(* PLC project GeneratedProgram, SafePLC-Gen SafePLC-Gen Multimodal 1.0 *)
(* stored: creationDateTime 2026-04-25T12:02:49.071447Z *)

PROGRAM GeneratedProgram
  VAR
    FirstScan : BOOL;
    TI_2909_Scaled : REAL;
    TT_2909_Scaled : REAL;
    TT_2911_Scaled : REAL;
    TT_2917_Scaled : REAL;
    TI_2917_Scaled : REAL;
    XI_2901A_Scaled : REAL;
    XI_2901B_Scaled : REAL;
    TI_2909_HH_SP : REAL;
    TI_2909_H_SP : REAL;
    TI_2909_L_SP : REAL;
    TI_2909_LL_SP : REAL;
    TI_2909_Deadband : REAL;
    TI_2909_HH_Latch : BOOL;
    TI_2909_LL_Latch : BOOL;
    TI_2909_HH : BOOL;
    TI_2909_H : BOOL;
    TI_2909_L : BOOL;
    TI_2909_LL : BOOL;
    TI_2909_HH_Ack : BOOL;
    TI_2909_LL_Ack : BOOL;
    TT_2909_HH_SP : REAL;
    TT_2909_H_SP : REAL;
    TT_2909_L_SP : REAL;
    TT_2909_LL_SP : REAL;
    TT_2909_Deadband : REAL;
    TT_2909_HH_Latch : BOOL;
    TT_2909_LL_Latch : BOOL;
    TT_2909_HH : BOOL;
    TT_2909_H : BOOL;
    TT_2909_L : BOOL;
    TT_2909_LL : BOOL;
    TT_2909_HH_Ack : BOOL;
    TT_2909_LL_Ack : BOOL;
    TT_2911_HH_SP : REAL;
    TT_2911_H_SP : REAL;
    TT_2911_L_SP : REAL;
    TT_2911_LL_SP : REAL;
    TT_2911_Deadband : REAL;
    TT_2911_HH_Latch : BOOL;
    TT_2911_LL_Latch : BOOL;
    TT_2911_HH : BOOL;
    TT_2911_H : BOOL;
    TT_2911_L : BOOL;
    TT_2911_LL : BOOL;
    TT_2911_HH_Ack : BOOL;
    TT_2911_LL_Ack : BOOL;
    TT_2917_HH_SP : REAL;
    TT_2917_H_SP : REAL;
    TT_2917_L_SP : REAL;
    TT_2917_LL_SP : REAL;
    TT_2917_Deadband : REAL;
    TT_2917_HH_Latch : BOOL;
    TT_2917_LL_Latch : BOOL;
    TT_2917_HH : BOOL;
    TT_2917_H : BOOL;
    TT_2917_L : BOOL;
    TT_2917_LL : BOOL;
    TT_2917_HH_Ack : BOOL;
    TT_2917_LL_Ack : BOOL;
    TI_2917_HH_SP : REAL;
    TI_2917_H_SP : REAL;
    TI_2917_L_SP : REAL;
    TI_2917_LL_SP : REAL;
    TI_2917_Deadband : REAL;
    TI_2917_HH_Latch : BOOL;
    TI_2917_LL_Latch : BOOL;
    TI_2917_HH : BOOL;
    TI_2917_H : BOOL;
    TI_2917_L : BOOL;
    TI_2917_LL : BOOL;
    TI_2917_HH_Ack : BOOL;
    TI_2917_LL_Ack : BOOL;
    XI_2901A_HH_SP : REAL;
    XI_2901A_H_SP : REAL;
    XI_2901A_L_SP : REAL;
    XI_2901A_LL_SP : REAL;
    XI_2901A_Deadband : REAL;
    XI_2901A_HH_Latch : BOOL;
    XI_2901A_LL_Latch : BOOL;
    XI_2901A_HH : BOOL;
    XI_2901A_H : BOOL;
    XI_2901A_L : BOOL;
    XI_2901A_LL : BOOL;
    XI_2901A_HH_Ack : BOOL;
    XI_2901A_LL_Ack : BOOL;
    XI_2901B_HH_SP : REAL;
    XI_2901B_H_SP : REAL;
    XI_2901B_L_SP : REAL;
    XI_2901B_LL_SP : REAL;
    XI_2901B_Deadband : REAL;
    XI_2901B_HH_Latch : BOOL;
    XI_2901B_LL_Latch : BOOL;
    XI_2901B_HH : BOOL;
    XI_2901B_H : BOOL;
    XI_2901B_L : BOOL;
    XI_2901B_LL : BOOL;
    XI_2901B_HH_Ack : BOOL;
    XI_2901B_LL_Ack : BOOL;
    LOOP_2917_TRIP : BOOL;
    LOOP_2901A_TRIP : BOOL;
    LOOP_2901B_TRIP : BOOL;
    VSHH_2901A_HH : BOOL;
    VSHH_2901A_LL : BOOL;
    VSHH_2901B_HH : BOOL;
    VSHH_2901B_LL : BOOL;
    SAFE_STATE : BOOL;
    MCC_A_Run : BOOL;
    MCC_B_Run : BOOL;
    MCC_A_Out : BOOL;
    MCC_B_Out : BOOL;
    Drive_A_SP : REAL;
    Drive_B_SP : REAL;
    Drive_A_Kp : REAL;
    Drive_A_Ki : REAL;
    Drive_B_Kp : REAL;
    Drive_B_Ki : REAL;
    Drive_A_Error : REAL;
    Drive_B_Error : REAL;
    Drive_A_Integral : REAL;
    Drive_B_Integral : REAL;
    Drive_A_Output : REAL;
    Drive_B_Output : REAL;
    StartDelay_A : TON;
    StartDelay_B : TON;
    RS_2901_Inlet_A_Upper : BOOL;
    RS_2901_Inlet_A_Lower : BOOL;
    RS_2901_Outlet_B_Upper : BOOL;
    RS_2901_Outlet_B_Lower : BOOL;
    BV_Inlet_A_Upper_1 : BOOL;
    BV_Inlet_A_Upper_2 : BOOL;
    BV_Inlet_A_Lower_1 : BOOL;
    BV_Inlet_A_Lower_2 : BOOL;
    BV_Outlet_B_Upper_1 : BOOL;
    BV_Outlet_B_Upper_2 : BOOL;
    BV_Outlet_B_Lower_1 : BOOL;
    BV_Outlet_B_Lower_2 : BOOL;
    CV_HY_2903A_1 : BOOL;
    CV_HY_2903A_2 : BOOL;
    CV_HY_2903B_1 : BOOL;
    CV_HY_2903B_2 : BOOL;
    CSO_Inlet_1 : BOOL;
    CSO_Inlet_2 : BOOL;
    FLV_Inlet : BOOL;
    BV_1IN_Drain : BOOL;
    Breather_A_8IN : BOOL;
    Breather_B_8IN : BOOL;
    NC_Valve_Outlet : BOOL;
    System_Alarm : BOOL;
  END_VAR

            IF FirstScan THEN
    LOOP_2917_TRIP          := TRUE;
    LOOP_2901A_TRIP         := TRUE;
    LOOP_2901B_TRIP         := TRUE;
    SAFE_STATE              := TRUE;
    MCC_A_Out               := FALSE;
    MCC_B_Out               := FALSE;
    MCC_A_Run               := FALSE;
    MCC_B_Run               := FALSE;
    HY_2903A_Out            := 6554;
    HY_2903B_Out            := 6554;
    KV_2904                 := FALSE;
    XL_2901A                := FALSE;
    XL_2901B                := FALSE;
    XA_2901A                := FALSE;
    XA_2901B                := FALSE;
    TI_2909_HH_Latch        := FALSE;
    TI_2909_LL_Latch        := FALSE;
    TT_2909_HH_Latch        := FALSE;
    TT_2909_LL_Latch        := FALSE;
    TT_2911_HH_Latch        := FALSE;
    TT_2911_LL_Latch        := FALSE;
    TT_2917_HH_Latch        := FALSE;
    TT_2917_LL_Latch        := FALSE;
    TI_2917_HH_Latch        := FALSE;
    TI_2917_LL_Latch        := FALSE;
    XI_2901A_HH_Latch       := FALSE;
    XI_2901A_LL_Latch       := FALSE;
    XI_2901B_HH_Latch       := FALSE;
    XI_2901B_LL_Latch       := FALSE;
    Drive_A_Integral        := 0.0;
    Drive_B_Integral        := 0.0;
    BV_1IN_Drain            := TRUE;
    StartDelay_A(IN := FALSE, PT := T#3S);
    StartDelay_B(IN := FALSE, PT := T#3S);
    FirstScan               := FALSE;
    RETURN;
END_IF;

TI_2909_Scaled  := ((INT_TO_REAL(TI_2909_Raw)  - 6554.0) / (32767.0 - 6554.0)) * 150.0;
TT_2909_Scaled  := ((INT_TO_REAL(TT_2909_Raw)  - 6554.0) / (32767.0 - 6554.0)) * 150.0;
TT_2911_Scaled  := ((INT_TO_REAL(TT_2911_Raw)  - 6554.0) / (32767.0 - 6554.0)) * 150.0;
TT_2917_Scaled  := ((INT_TO_REAL(TT_2917_Raw)  - 6554.0) / (32767.0 - 6554.0)) * 150.0;
TI_2917_Scaled  := ((INT_TO_REAL(TI_2917_Raw)  - 6554.0) / (32767.0 - 6554.0)) * 150.0;
XI_2901A_Scaled := ((INT_TO_REAL(XI_2901A_Raw) - 6554.0) / (32767.0 - 6554.0)) * 100.0;
XI_2901B_Scaled := ((INT_TO_REAL(XI_2901B_Raw) - 6554.0) / (32767.0 - 6554.0)) * 100.0;

IF TI_2909_Scaled >= TI_2909_HH_SP THEN
    TI_2909_HH_Latch := TRUE;
ELSIF TI_2909_Scaled <= (TI_2909_HH_SP - TI_2909_Deadband) AND TI_2909_HH_Ack THEN
    TI_2909_HH_Latch := FALSE;
END_IF;
TI_2909_HH := TI_2909_HH_Latch;
TI_2909_H  := TI_2909_Scaled >= TI_2909_H_SP;
TI_2909_L  := TI_2909_Scaled <= TI_2909_L_SP;
IF TI_2909_Scaled <= TI_2909_LL_SP THEN
    TI_2909_LL_Latch := TRUE;
ELSIF TI_2909_Scaled >= (TI_2909_LL_SP + TI_2909_Deadband) AND TI_2909_LL_Ack THEN
    TI_2909_LL_Latch := FALSE;
END_IF;
TI_2909_LL := TI_2909_LL_Latch;

IF TT_2909_Scaled >= TT_2909_HH_SP THEN
    TT_2909_HH_Latch := TRUE;
ELSIF TT_2909_Scaled <= (TT_2909_HH_SP - TT_2909_Deadband) AND TT_2909_HH_Ack THEN
    TT_2909_HH_Latch := FALSE;
END_IF;
TT_2909_HH := TT_2909_HH_Latch;
TT_2909_H  := TT_2909_Scaled >= TT_2909_H_SP;
TT_2909_L  := TT_2909_Scaled <= TT_2909_L_SP;
IF TT_2909_Scaled <= TT_2909_LL_SP THEN
    TT_2909_LL_Latch := TRUE;
ELSIF TT_2909_Scaled >= (TT_2909_LL_SP + TT_2909_Deadband) AND TT_2909_LL_Ack THEN
    TT_2909_LL_Latch := FALSE;
END_IF;
TT_2909_LL := TT_2909_LL_Latch;

IF TT_2911_Scaled >= TT_2911_HH_SP THEN
    TT_2911_HH_Latch := TRUE;
ELSIF TT_2911_Scaled <= (TT_2911_HH_SP - TT_2911_Deadband) AND TT_2911_HH_Ack THEN
    TT_2911_HH_Latch := FALSE;
END_IF;
TT_2911_HH := TT_2911_HH_Latch;
TT_2911_H  := TT_2911_Scaled >= TT_2911_H_SP;
TT_2911_L  := TT_2911_Scaled <= TT_2911_L_SP;
IF TT_2911_Scaled <= TT_2911_LL_SP THEN
    TT_2911_LL_Latch := TRUE;
ELSIF TT_2911_Scaled >= (TT_2911_LL_SP + TT_2911_Deadband) AND TT_2911_LL_Ack THEN
    TT_2911_LL_Latch := FALSE;
END_IF;
TT_2911_LL := TT_2911_LL_Latch;

IF TT_2917_Scaled >= TT_2917_HH_SP THEN
    TT_2917_HH_Latch := TRUE;
ELSIF TT_2917_Scaled <= (TT_2917_HH_SP - TT_2917_Deadband) AND TT_2917_HH_Ack THEN
    TT_2917_HH_Latch := FALSE;
END_IF;
TT_2917_HH := TT_2917_HH_Latch;
TT_2917_H  := TT_2917_Scaled >= TT_2917_H_SP;
TT_2917_L  := TT_2917_Scaled <= TT_2917_L_SP;
IF TT_2917_Scaled <= TT_2917_LL_SP THEN
    TT_2917_LL_Latch := TRUE;
ELSIF TT_2917_Scaled >= (TT_2917_LL_SP + TT_2917_Deadband) AND TT_2917_LL_Ack THEN
    TT_2917_LL_Latch := FALSE;
END_IF;
TT_2917_LL := TT_2917_LL_Latch;

IF TI_2917_Scaled >= TI_2917_HH_SP THEN
    TI_2917_HH_Latch := TRUE;
ELSIF TI_2917_Scaled <= (TI_2917_HH_SP - TI_2917_Deadband) AND TI_2917_HH_Ack THEN
    TI_2917_HH_Latch := FALSE;
END_IF;
TI_2917_HH := TI_2917_HH_Latch;
TI_2917_H  := TI_2917_Scaled >= TI_2917_H_SP;
TI_2917_L  := TI_2917_Scaled <= TI_2917_L_SP;
IF TI_2917_Scaled <= TI_2917_LL_SP THEN
    TI_2917_LL_Latch := TRUE;
ELSIF TI_2917_Scaled >= (TI_2917_LL_SP + TI_2917_Deadband) AND TI_2917_LL_Ack THEN
    TI_2917_LL_Latch := FALSE;
END_IF;
TI_2917_LL := TI_2917_LL_Latch;

IF XI_2901A_Scaled >= XI_2901A_HH_SP THEN
    XI_2901A_HH_Latch := TRUE;
ELSIF XI_2901A_Scaled <= (XI_2901A_HH_SP - XI_2901A_Deadband) AND XI_2901A_HH_Ack THEN
    XI_2901A_HH_Latch := FALSE;
END_IF;
XI_2901A_HH := XI_2901A_HH_Latch;
XI_2901A_H  := XI_2901A_Scaled >= XI_2901A_H_SP;
XI_2901A_L  := XI_2901A_Scaled <= XI_2901A_L_SP;
IF XI_2901A_Scaled <= XI_2901A_LL_SP THEN
    XI_2901A_LL_Latch := TRUE;
ELSIF XI_2901A_Scaled >= (XI_2901A_LL_SP + XI_2901A_Deadband) AND XI_2901A_LL_Ack THEN
    XI_2901A_LL_Latch := FALSE;
END_IF;
XI_2901A_LL := XI_2901A_LL_Latch;

IF XI_2901B_Scaled >= XI_2901B_HH_SP THEN
    XI_2901B_HH_Latch := TRUE;
ELSIF XI_2901B_Scaled <= (XI_2901B_HH_SP - XI_2901B_Deadband) AND XI_2901B_HH_Ack THEN
    XI_2901B_HH_Latch := FALSE;
END_IF;
XI_2901B_HH := XI_2901B_HH_Latch;
XI_2901B_H  := XI_2901B_Scaled >= XI_2901B_H_SP;
XI_2901B_L  := XI_2901B_Scaled <= XI_2901B_L_SP;
IF XI_2901B_Scaled <= XI_2901B_LL_SP THEN
    XI_2901B_LL_Latch := TRUE;
ELSIF XI_2901B_Scaled >= (XI_2901B_LL_SP + XI_2901B_Deadband) AND XI_2901B_LL_Ack THEN
    XI_2901B_LL_Latch := FALSE;
END_IF;
XI_2901B_LL := XI_2901B_LL_Latch;

VSHH_2901A_HH := VSHH_2901A;
VSHH_2901A_LL := FALSE;
VSHH_2901B_HH := VSHH_2901B;
VSHH_2901B_LL := FALSE;

IF TT_2917_HH OR TT_2917_LL OR TI_2917_HH OR TI_2917_LL OR PSD_2917 THEN
    LOOP_2917_TRIP := TRUE;
ELSIF LOOP_2917_TRIP AND MANUAL_RESET
      AND NOT TT_2917_HH AND NOT TT_2917_LL
      AND NOT TI_2917_HH AND NOT TI_2917_LL
      AND NOT PSD_2917 THEN
    LOOP_2917_TRIP := FALSE;
END_IF;

IF VSHH_2901A_HH OR VSHH_2901A_LL THEN
    LOOP_2901A_TRIP := TRUE;
ELSIF LOOP_2901A_TRIP AND MANUAL_RESET
      AND NOT VSHH_2901A_HH AND NOT VSHH_2901A_LL THEN
    LOOP_2901A_TRIP := FALSE;
END_IF;

IF VSHH_2901B_HH OR VSHH_2901B_LL THEN
    LOOP_2901B_TRIP := TRUE;
ELSIF LOOP_2901B_TRIP AND MANUAL_RESET
      AND NOT VSHH_2901B_HH AND NOT VSHH_2901B_LL THEN
    LOOP_2901B_TRIP := FALSE;
END_IF;

SAFE_STATE := ESTOP OR ESD_3200
              OR HS_EMGSTOP_A_2901A OR HS_EMGSTOP_B_2901B
              OR LOOP_2917_TRIP OR LOOP_2901A_TRIP OR LOOP_2901B_TRIP;

StartDelay_A(IN := MCC_A_Run AND NOT SAFE_STATE, PT := T#3S);
StartDelay_B(IN := MCC_B_Run AND NOT SAFE_STATE, PT := T#3S);

IF NOT SAFE_STATE THEN
    IF HS_2901A1 THEN
        IF HS_START_STOP_A_2901A THEN
            MCC_A_Run := TRUE;
        ELSIF NOT HS_2901A THEN
            MCC_A_Run := FALSE;
        END_IF;
    ELSE
        MCC_A_Run := HS_2901A2;
    END_IF;

    MCC_A_Out := StartDelay_A.Q;

    IF MCC_A_Out THEN
        Drive_A_Error    := Drive_A_SP - XI_2901A_Scaled;
        Drive_A_Integral := Drive_A_Integral + (Drive_A_Ki * Drive_A_Error);
        IF Drive_A_Integral > 100.0 THEN
            Drive_A_Integral := 100.0;
        ELSIF Drive_A_Integral < 0.0 THEN
            Drive_A_Integral := 0.0;
        END_IF;
        Drive_A_Output := (Drive_A_Kp * Drive_A_Error) + Drive_A_Integral;
        IF Drive_A_Output > 100.0 THEN
            Drive_A_Output := 100.0;
        ELSIF Drive_A_Output < 0.0 THEN
            Drive_A_Output := 0.0;
        END_IF;
        HY_2903A_Out := REAL_TO_INT(6554.0 + (Drive_A_Output / 100.0) * (32767.0 - 6554.0));
    ELSE
        HY_2903A_Out     := 6554;
        Drive_A_Integral := 0.0;
    END_IF;

    IF HS_2901B1 THEN
        IF HS_START_STOP_B_2901B THEN
            MCC_B_Run := TRUE;
        ELSIF NOT HS_2901B THEN
            MCC_B_Run := FALSE;
        END_IF;
    ELSE
        MCC_B_Run := HS_2901B2;
    END_IF;

    MCC_B_Out := StartDelay_B.Q;

    IF MCC_B_Out THEN
        Drive_B_Error    := Drive_B_SP - XI_2901B_Scaled;
        Drive_B_Integral := Drive_B_Integral + (Drive_B_Ki * Drive_B_Error);
        IF Drive_B_Integral > 100.0 THEN
            Drive_B_Integral := 100.0;
        ELSIF Drive_B_Integral < 0.0 THEN
            Drive_B_Integral := 0.0;
        END_IF;
        Drive_B_Output := (Drive_B_Kp * Drive_B_Error) + Drive_B_Integral;
        IF Drive_B_Output > 100.0 THEN
            Drive_B_Output := 100.0;
        ELSIF Drive_B_Output < 0.0 THEN
            Drive_B_Output := 0.0;
        END_IF;
        HY_2903B_Out := REAL_TO_INT(6554.0 + (Drive_B_Output / 100.0) * (32767.0 - 6554.0));
    ELSE
        HY_2903B_Out     := 6554;
        Drive_B_Integral := 0.0;
    END_IF;

    KV_2904                := MCC_A_Out OR MCC_B_Out;
    RS_2901_Inlet_A_Upper  := MCC_A_Out;
    RS_2901_Inlet_A_Lower  := MCC_A_Out;
    RS_2901_Outlet_B_Upper := MCC_B_Out;
    RS_2901_Outlet_B_Lower := MCC_B_Out;
    BV_Inlet_A_Upper_1     := MCC_A_Out;
    BV_Inlet_A_Upper_2     := MCC_A_Out;
    BV_Inlet_A_Lower_1     := MCC_A_Out;
    BV_Inlet_A_Lower_2     := MCC_A_Out;
    BV_Outlet_B_Upper_1    := MCC_B_Out;
    BV_Outlet_B_Upper_2    := MCC_B_Out;
    BV_Outlet_B_Lower_1    := MCC_B_Out;
    BV_Outlet_B_Lower_2    := MCC_B_Out;
    CV_HY_2903A_1          := MCC_A_Out;
    CV_HY_2903A_2          := MCC_A_Out;
    CV_HY_2903B_1          := MCC_B_Out;
    CV_HY_2903B_2          := MCC_B_Out;
    CSO_Inlet_1            := MCC_A_Out OR MCC_B_Out;
    CSO_Inlet_2            := MCC_A_Out OR MCC_B_Out;
    FLV_Inlet              := MCC_A_Out OR MCC_B_Out;
    BV_1IN_Drain           := NOT (MCC_A_Out OR MCC_B_Out);
    Breather_A_8IN         := MCC_A_Out;
    Breather_B_8IN         := MCC_B_Out;
    NC_Valve_Outlet        := MCC_A_Out OR MCC_B_Out;
    XL_2901A               := MCC_A_Out;
    XL_2901B               := MCC_B_Out;
    XA_2901A               := LOOP_2901A_TRIP OR XI_2901A_HH;
    XA_2901B               := LOOP_2901B_TRIP OR XI_2901B_HH;
ELSE
    MCC_A_Out              := FALSE;
    MCC_B_Out              := FALSE;
    MCC_A_Run              := FALSE;
    MCC_B_Run              := FALSE;
    HY_2903A_Out           := 6554;
    HY_2903B_Out           := 6554;
    KV_2904                := FALSE;
    XL_2901A               := FALSE;
    XL_2901B               := FALSE;
    XA_2901A               := TRUE;
    XA_2901B               := TRUE;
    Drive_A_Integral       := 0.0;
    Drive_B_Integral       := 0.0;
    RS_2901_Inlet_A_Upper  := FALSE;
    RS_2901_Inlet_A_Lower  := FALSE;
    RS_2901_Outlet_B_Upper := FALSE;
    RS_2901_Outlet_B_Lower := FALSE;
    BV_Inlet_A_Upper_1     := FALSE;
    BV_Inlet_A_Upper_2     := FALSE;
    BV_Inlet_A_Lower_1     := FALSE;
    BV_Inlet_A_Lower_2     := FALSE;
    BV_Outlet_B_Upper_1    := FALSE;
    BV_Outlet_B_Upper_2    := FALSE;
    BV_Outlet_B_Lower_1    := FALSE;
    BV_Outlet_B_Lower_2    := FALSE;
    CV_HY_2903A_1          := FALSE;
    CV_HY_2903A_2          := FALSE;
    CV_HY_2903B_1          := FALSE;
    CV_HY_2903B_2          := FALSE;
    CSO_Inlet_1            := FALSE;
    CSO_Inlet_2            := FALSE;
    FLV_Inlet              := FALSE;
    BV_1IN_Drain           := TRUE;
    Breather_A_8IN         := FALSE;
    Breather_B_8IN         := FALSE;
    NC_Valve_Outlet        := FALSE;
END_IF;

System_Alarm :=
    TI_2909_HH_Latch  OR TI_2909_LL_Latch  OR TI_2909_H  OR TI_2909_L  OR
    TT_2909_HH_Latch  OR TT_2909_LL_Latch  OR TT_2909_H  OR TT_2909_L  OR
    TT_2911_HH_Latch  OR TT_2911_LL_Latch  OR TT_2911_H  OR TT_2911_L  OR
    TT_2917_HH_Latch  OR TT_2917_LL_Latch  OR TT_2917_H  OR TT_2917_L  OR
    TI_2917_HH_Latch  OR TI_2917_LL_Latch  OR TI_2917_H  OR TI_2917_L  OR
    XI_2901A_HH_Latch OR XI_2901A_LL_Latch OR XI_2901A_H OR XI_2901A_L OR
    XI_2901B_HH_Latch OR XI_2901B_LL_Latch OR XI_2901B_H OR XI_2901B_L OR
    LOOP_2917_TRIP OR LOOP_2901A_TRIP OR LOOP_2901B_TRIP OR SAFE_STATE;
          
END_PROGRAM

CONFIGURATION Config0
  RESOURCE Res0 ON PLC
    TASK MainTask(INTERVAL := T#20ms, PRIORITY := 0);
    PROGRAM Main : GeneratedProgram;
  END_RESOURCE
END_CONFIGURATION
